Fanuc KAREL source: KA00028.KL

PROGRAM KA00028
%NOLOCKGROUP
VAR
  SRC: BOOLEAN
  DST: STRING[80]
BEGIN
  SRC = TRUE
  DST = SRC
END KA00028
